(* IEC 61131-3 sources: STAR-PLC-Agent/results/raw/codex_matrix_resume_20261114/codex_deepseek/SELF004/functional/attempt_0001, 1 file *)

(* ---- test_program.st ---- *)
PROGRAM PLC_PRG
VAR
 BenchStep : UDINT := 0;
 BenchCalls : UDINT := 0;
 BenchDone : BOOL := FALSE;
 BenchUut0 : FB_Task;
 BenchUut1 : FB_Task;
 BenchUut2 : FB_Task;
 BenchUut3 : FB_Task;
 BenchUut4 : FB_Task;
 BenchUut5 : FB_Task;
 BenchUut6 : FB_Task;
 BenchUut7 : FB_Task;
 BenchUut8 : FB_Task;
 TraceIn_Start : ARRAY[0..60] OF BOOL;
 TraceIn_Stop : ARRAY[0..60] OF BOOL;
 TraceIn_AtExit : ARRAY[0..60] OF BOOL;
 TraceIn_Jam : ARRAY[0..60] OF BOOL;
 TraceIn_Reset : ARRAY[0..60] OF BOOL;
 TraceOut_Belt : ARRAY[0..60] OF BOOL;
 TraceOut_Complete : ARRAY[0..60] OF BOOL;
 TraceOut_Fault : ARRAY[0..60] OF BOOL;
END_VAR

IF NOT BenchDone THEN
 CASE BenchStep OF
 0:
   BenchUut0.Start := TRUE;
   BenchUut0.Stop := FALSE;
   BenchUut0.AtExit := FALSE;
   BenchUut0.Jam := FALSE;
   BenchUut0.Reset := FALSE;
   TraceIn_Start[0] := BenchUut0.Start;
   TraceIn_Stop[0] := BenchUut0.Stop;
   TraceIn_AtExit[0] := BenchUut0.AtExit;
   TraceIn_Jam[0] := BenchUut0.Jam;
   TraceIn_Reset[0] := BenchUut0.Reset;
   BenchUut0();
   TraceOut_Belt[0] := BenchUut0.Belt;
   TraceOut_Complete[0] := BenchUut0.Complete;
   TraceOut_Fault[0] := BenchUut0.Fault;
   BenchCalls := BenchCalls + 1;
 1:
   BenchUut0.Start := FALSE;
   BenchUut0.Stop := FALSE;
   BenchUut0.AtExit := FALSE;
   BenchUut0.Jam := FALSE;
   BenchUut0.Reset := FALSE;
   TraceIn_Start[1] := BenchUut0.Start;
   TraceIn_Stop[1] := BenchUut0.Stop;
   TraceIn_AtExit[1] := BenchUut0.AtExit;
   TraceIn_Jam[1] := BenchUut0.Jam;
   TraceIn_Reset[1] := BenchUut0.Reset;
   BenchUut0();
   TraceOut_Belt[1] := BenchUut0.Belt;
   TraceOut_Complete[1] := BenchUut0.Complete;
   TraceOut_Fault[1] := BenchUut0.Fault;
   BenchCalls := BenchCalls + 1;
 2:
   BenchUut0.Start := FALSE;
   BenchUut0.Stop := FALSE;
   BenchUut0.AtExit := TRUE;
   BenchUut0.Jam := FALSE;
   BenchUut0.Reset := FALSE;
   TraceIn_Start[2] := BenchUut0.Start;
   TraceIn_Stop[2] := BenchUut0.Stop;
   TraceIn_AtExit[2] := BenchUut0.AtExit;
   TraceIn_Jam[2] := BenchUut0.Jam;
   TraceIn_Reset[2] := BenchUut0.Reset;
   BenchUut0();
   TraceOut_Belt[2] := BenchUut0.Belt;
   TraceOut_Complete[2] := BenchUut0.Complete;
   TraceOut_Fault[2] := BenchUut0.Fault;
   BenchCalls := BenchCalls + 1;
 3:
   BenchUut0.Start := TRUE;
   BenchUut0.Stop := FALSE;
   BenchUut0.AtExit := FALSE;
   BenchUut0.Jam := FALSE;
   BenchUut0.Reset := FALSE;
   TraceIn_Start[3] := BenchUut0.Start;
   TraceIn_Stop[3] := BenchUut0.Stop;
   TraceIn_AtExit[3] := BenchUut0.AtExit;
   TraceIn_Jam[3] := BenchUut0.Jam;
   TraceIn_Reset[3] := BenchUut0.Reset;
   BenchUut0();
   TraceOut_Belt[3] := BenchUut0.Belt;
   TraceOut_Complete[3] := BenchUut0.Complete;
   TraceOut_Fault[3] := BenchUut0.Fault;
   BenchCalls := BenchCalls + 1;
 4:
   BenchUut0.Start := FALSE;
   BenchUut0.Stop := FALSE;
   BenchUut0.AtExit := FALSE;
   BenchUut0.Jam := FALSE;
   BenchUut0.Reset := TRUE;
   TraceIn_Start[4] := BenchUut0.Start;
   TraceIn_Stop[4] := BenchUut0.Stop;
   TraceIn_AtExit[4] := BenchUut0.AtExit;
   TraceIn_Jam[4] := BenchUut0.Jam;
   TraceIn_Reset[4] := BenchUut0.Reset;
   BenchUut0();
   TraceOut_Belt[4] := BenchUut0.Belt;
   TraceOut_Complete[4] := BenchUut0.Complete;
   TraceOut_Fault[4] := BenchUut0.Fault;
   BenchCalls := BenchCalls + 1;
 5:
   BenchUut1.Start := TRUE;
   BenchUut1.Stop := FALSE;
   BenchUut1.AtExit := FALSE;
   BenchUut1.Jam := FALSE;
   BenchUut1.Reset := FALSE;
   TraceIn_Start[5] := BenchUut1.Start;
   TraceIn_Stop[5] := BenchUut1.Stop;
   TraceIn_AtExit[5] := BenchUut1.AtExit;
   TraceIn_Jam[5] := BenchUut1.Jam;
   TraceIn_Reset[5] := BenchUut1.Reset;
   BenchUut1();
   TraceOut_Belt[5] := BenchUut1.Belt;
   TraceOut_Complete[5] := BenchUut1.Complete;
   TraceOut_Fault[5] := BenchUut1.Fault;
   BenchCalls := BenchCalls + 1;
 6:
   BenchUut1.Start := TRUE;
   BenchUut1.Stop := FALSE;
   BenchUut1.AtExit := FALSE;
   BenchUut1.Jam := TRUE;
   BenchUut1.Reset := TRUE;
   TraceIn_Start[6] := BenchUut1.Start;
   TraceIn_Stop[6] := BenchUut1.Stop;
   TraceIn_AtExit[6] := BenchUut1.AtExit;
   TraceIn_Jam[6] := BenchUut1.Jam;
   TraceIn_Reset[6] := BenchUut1.Reset;
   BenchUut1();
   TraceOut_Belt[6] := BenchUut1.Belt;
   TraceOut_Complete[6] := BenchUut1.Complete;
   TraceOut_Fault[6] := BenchUut1.Fault;
   BenchCalls := BenchCalls + 1;
 7:
   BenchUut1.Start := TRUE;
   BenchUut1.Stop := FALSE;
   BenchUut1.AtExit := FALSE;
   BenchUut1.Jam := FALSE;
   BenchUut1.Reset := FALSE;
   TraceIn_Start[7] := BenchUut1.Start;
   TraceIn_Stop[7] := BenchUut1.Stop;
   TraceIn_AtExit[7] := BenchUut1.AtExit;
   TraceIn_Jam[7] := BenchUut1.Jam;
   TraceIn_Reset[7] := BenchUut1.Reset;
   BenchUut1();
   TraceOut_Belt[7] := BenchUut1.Belt;
   TraceOut_Complete[7] := BenchUut1.Complete;
   TraceOut_Fault[7] := BenchUut1.Fault;
   BenchCalls := BenchCalls + 1;
 8:
   BenchUut1.Start := TRUE;
   BenchUut1.Stop := FALSE;
   BenchUut1.AtExit := FALSE;
   BenchUut1.Jam := FALSE;
   BenchUut1.Reset := TRUE;
   TraceIn_Start[8] := BenchUut1.Start;
   TraceIn_Stop[8] := BenchUut1.Stop;
   TraceIn_AtExit[8] := BenchUut1.AtExit;
   TraceIn_Jam[8] := BenchUut1.Jam;
   TraceIn_Reset[8] := BenchUut1.Reset;
   BenchUut1();
   TraceOut_Belt[8] := BenchUut1.Belt;
   TraceOut_Complete[8] := BenchUut1.Complete;
   TraceOut_Fault[8] := BenchUut1.Fault;
   BenchCalls := BenchCalls + 1;
 9:
   BenchUut1.Start := TRUE;
   BenchUut1.Stop := FALSE;
   BenchUut1.AtExit := TRUE;
   BenchUut1.Jam := FALSE;
   BenchUut1.Reset := FALSE;
   TraceIn_Start[9] := BenchUut1.Start;
   TraceIn_Stop[9] := BenchUut1.Stop;
   TraceIn_AtExit[9] := BenchUut1.AtExit;
   TraceIn_Jam[9] := BenchUut1.Jam;
   TraceIn_Reset[9] := BenchUut1.Reset;
   BenchUut1();
   TraceOut_Belt[9] := BenchUut1.Belt;
   TraceOut_Complete[9] := BenchUut1.Complete;
   TraceOut_Fault[9] := BenchUut1.Fault;
   BenchCalls := BenchCalls + 1;
 10:
   BenchUut1.Start := TRUE;
   BenchUut1.Stop := TRUE;
   BenchUut1.AtExit := FALSE;
   BenchUut1.Jam := FALSE;
   BenchUut1.Reset := FALSE;
   TraceIn_Start[10] := BenchUut1.Start;
   TraceIn_Stop[10] := BenchUut1.Stop;
   TraceIn_AtExit[10] := BenchUut1.AtExit;
   TraceIn_Jam[10] := BenchUut1.Jam;
   TraceIn_Reset[10] := BenchUut1.Reset;
   BenchUut1();
   TraceOut_Belt[10] := BenchUut1.Belt;
   TraceOut_Complete[10] := BenchUut1.Complete;
   TraceOut_Fault[10] := BenchUut1.Fault;
   BenchCalls := BenchCalls + 1;
 11:
   BenchUut2.Start := TRUE;
   BenchUut2.Stop := FALSE;
   BenchUut2.AtExit := FALSE;
   BenchUut2.Jam := FALSE;
   BenchUut2.Reset := FALSE;
   TraceIn_Start[11] := BenchUut2.Start;
   TraceIn_Stop[11] := BenchUut2.Stop;
   TraceIn_AtExit[11] := BenchUut2.AtExit;
   TraceIn_Jam[11] := BenchUut2.Jam;
   TraceIn_Reset[11] := BenchUut2.Reset;
   BenchUut2();
   TraceOut_Belt[11] := BenchUut2.Belt;
   TraceOut_Complete[11] := BenchUut2.Complete;
   TraceOut_Fault[11] := BenchUut2.Fault;
   BenchCalls := BenchCalls + 1;
 12:
   BenchUut2.Start := FALSE;
   BenchUut2.Stop := TRUE;
   BenchUut2.AtExit := TRUE;
   BenchUut2.Jam := FALSE;
   BenchUut2.Reset := FALSE;
   TraceIn_Start[12] := BenchUut2.Start;
   TraceIn_Stop[12] := BenchUut2.Stop;
   TraceIn_AtExit[12] := BenchUut2.AtExit;
   TraceIn_Jam[12] := BenchUut2.Jam;
   TraceIn_Reset[12] := BenchUut2.Reset;
   BenchUut2();
   TraceOut_Belt[12] := BenchUut2.Belt;
   TraceOut_Complete[12] := BenchUut2.Complete;
   TraceOut_Fault[12] := BenchUut2.Fault;
   BenchCalls := BenchCalls + 1;
 13:
   BenchUut2.Start := TRUE;
   BenchUut2.Stop := FALSE;
   BenchUut2.AtExit := FALSE;
   BenchUut2.Jam := FALSE;
   BenchUut2.Reset := FALSE;
   TraceIn_Start[13] := BenchUut2.Start;
   TraceIn_Stop[13] := BenchUut2.Stop;
   TraceIn_AtExit[13] := BenchUut2.AtExit;
   TraceIn_Jam[13] := BenchUut2.Jam;
   TraceIn_Reset[13] := BenchUut2.Reset;
   BenchUut2();
   TraceOut_Belt[13] := BenchUut2.Belt;
   TraceOut_Complete[13] := BenchUut2.Complete;
   TraceOut_Fault[13] := BenchUut2.Fault;
   BenchCalls := BenchCalls + 1;
 14:
   BenchUut2.Start := FALSE;
   BenchUut2.Stop := FALSE;
   BenchUut2.AtExit := FALSE;
   BenchUut2.Jam := FALSE;
   BenchUut2.Reset := TRUE;
   TraceIn_Start[14] := BenchUut2.Start;
   TraceIn_Stop[14] := BenchUut2.Stop;
   TraceIn_AtExit[14] := BenchUut2.AtExit;
   TraceIn_Jam[14] := BenchUut2.Jam;
   TraceIn_Reset[14] := BenchUut2.Reset;
   BenchUut2();
   TraceOut_Belt[14] := BenchUut2.Belt;
   TraceOut_Complete[14] := BenchUut2.Complete;
   TraceOut_Fault[14] := BenchUut2.Fault;
   BenchCalls := BenchCalls + 1;
 15:
   BenchUut2.Start := TRUE;
   BenchUut2.Stop := FALSE;
   BenchUut2.AtExit := FALSE;
   BenchUut2.Jam := FALSE;
   BenchUut2.Reset := FALSE;
   TraceIn_Start[15] := BenchUut2.Start;
   TraceIn_Stop[15] := BenchUut2.Stop;
   TraceIn_AtExit[15] := BenchUut2.AtExit;
   TraceIn_Jam[15] := BenchUut2.Jam;
   TraceIn_Reset[15] := BenchUut2.Reset;
   BenchUut2();
   TraceOut_Belt[15] := BenchUut2.Belt;
   TraceOut_Complete[15] := BenchUut2.Complete;
   TraceOut_Fault[15] := BenchUut2.Fault;
   BenchCalls := BenchCalls + 1;
 16:
   BenchUut2.Start := FALSE;
   BenchUut2.Stop := FALSE;
   BenchUut2.AtExit := TRUE;
   BenchUut2.Jam := FALSE;
   BenchUut2.Reset := FALSE;
   TraceIn_Start[16] := BenchUut2.Start;
   TraceIn_Stop[16] := BenchUut2.Stop;
   TraceIn_AtExit[16] := BenchUut2.AtExit;
   TraceIn_Jam[16] := BenchUut2.Jam;
   TraceIn_Reset[16] := BenchUut2.Reset;
   BenchUut2();
   TraceOut_Belt[16] := BenchUut2.Belt;
   TraceOut_Complete[16] := BenchUut2.Complete;
   TraceOut_Fault[16] := BenchUut2.Fault;
   BenchCalls := BenchCalls + 1;
 17:
   BenchUut2.Start := FALSE;
   BenchUut2.Stop := TRUE;
   BenchUut2.AtExit := TRUE;
   BenchUut2.Jam := FALSE;
   BenchUut2.Reset := FALSE;
   TraceIn_Start[17] := BenchUut2.Start;
   TraceIn_Stop[17] := BenchUut2.Stop;
   TraceIn_AtExit[17] := BenchUut2.AtExit;
   TraceIn_Jam[17] := BenchUut2.Jam;
   TraceIn_Reset[17] := BenchUut2.Reset;
   BenchUut2();
   TraceOut_Belt[17] := BenchUut2.Belt;
   TraceOut_Complete[17] := BenchUut2.Complete;
   TraceOut_Fault[17] := BenchUut2.Fault;
   BenchCalls := BenchCalls + 1;
 18:
   BenchUut2.Start := FALSE;
   BenchUut2.Stop := FALSE;
   BenchUut2.AtExit := FALSE;
   BenchUut2.Jam := TRUE;
   BenchUut2.Reset := FALSE;
   TraceIn_Start[18] := BenchUut2.Start;
   TraceIn_Stop[18] := BenchUut2.Stop;
   TraceIn_AtExit[18] := BenchUut2.AtExit;
   TraceIn_Jam[18] := BenchUut2.Jam;
   TraceIn_Reset[18] := BenchUut2.Reset;
   BenchUut2();
   TraceOut_Belt[18] := BenchUut2.Belt;
   TraceOut_Complete[18] := BenchUut2.Complete;
   TraceOut_Fault[18] := BenchUut2.Fault;
   BenchCalls := BenchCalls + 1;
 19:
   BenchUut2.Start := TRUE;
   BenchUut2.Stop := TRUE;
   BenchUut2.AtExit := FALSE;
   BenchUut2.Jam := FALSE;
   BenchUut2.Reset := FALSE;
   TraceIn_Start[19] := BenchUut2.Start;
   TraceIn_Stop[19] := BenchUut2.Stop;
   TraceIn_AtExit[19] := BenchUut2.AtExit;
   TraceIn_Jam[19] := BenchUut2.Jam;
   TraceIn_Reset[19] := BenchUut2.Reset;
   BenchUut2();
   TraceOut_Belt[19] := BenchUut2.Belt;
   TraceOut_Complete[19] := BenchUut2.Complete;
   TraceOut_Fault[19] := BenchUut2.Fault;
   BenchCalls := BenchCalls + 1;
 20:
   BenchUut2.Start := FALSE;
   BenchUut2.Stop := FALSE;
   BenchUut2.AtExit := FALSE;
   BenchUut2.Jam := FALSE;
   BenchUut2.Reset := TRUE;
   TraceIn_Start[20] := BenchUut2.Start;
   TraceIn_Stop[20] := BenchUut2.Stop;
   TraceIn_AtExit[20] := BenchUut2.AtExit;
   TraceIn_Jam[20] := BenchUut2.Jam;
   TraceIn_Reset[20] := BenchUut2.Reset;
   BenchUut2();
   TraceOut_Belt[20] := BenchUut2.Belt;
   TraceOut_Complete[20] := BenchUut2.Complete;
   TraceOut_Fault[20] := BenchUut2.Fault;
   BenchCalls := BenchCalls + 1;
 21:
   BenchUut3.Start := TRUE;
   BenchUut3.Stop := FALSE;
   BenchUut3.AtExit := FALSE;
   BenchUut3.Jam := FALSE;
   BenchUut3.Reset := FALSE;
   TraceIn_Start[21] := BenchUut3.Start;
   TraceIn_Stop[21] := BenchUut3.Stop;
   TraceIn_AtExit[21] := BenchUut3.AtExit;
   TraceIn_Jam[21] := BenchUut3.Jam;
   TraceIn_Reset[21] := BenchUut3.Reset;
   BenchUut3();
   TraceOut_Belt[21] := BenchUut3.Belt;
   TraceOut_Complete[21] := BenchUut3.Complete;
   TraceOut_Fault[21] := BenchUut3.Fault;
   BenchCalls := BenchCalls + 1;
 22:
   BenchUut3.Start := FALSE;
   BenchUut3.Stop := FALSE;
   BenchUut3.AtExit := FALSE;
   BenchUut3.Jam := FALSE;
   BenchUut3.Reset := FALSE;
   TraceIn_Start[22] := BenchUut3.Start;
   TraceIn_Stop[22] := BenchUut3.Stop;
   TraceIn_AtExit[22] := BenchUut3.AtExit;
   TraceIn_Jam[22] := BenchUut3.Jam;
   TraceIn_Reset[22] := BenchUut3.Reset;
   BenchUut3();
   TraceOut_Belt[22] := BenchUut3.Belt;
   TraceOut_Complete[22] := BenchUut3.Complete;
   TraceOut_Fault[22] := BenchUut3.Fault;
   BenchCalls := BenchCalls + 1;
 23:
   BenchUut3.Start := FALSE;
   BenchUut3.Stop := FALSE;
   BenchUut3.AtExit := TRUE;
   BenchUut3.Jam := FALSE;
   BenchUut3.Reset := FALSE;
   TraceIn_Start[23] := BenchUut3.Start;
   TraceIn_Stop[23] := BenchUut3.Stop;
   TraceIn_AtExit[23] := BenchUut3.AtExit;
   TraceIn_Jam[23] := BenchUut3.Jam;
   TraceIn_Reset[23] := BenchUut3.Reset;
   BenchUut3();
   TraceOut_Belt[23] := BenchUut3.Belt;
   TraceOut_Complete[23] := BenchUut3.Complete;
   TraceOut_Fault[23] := BenchUut3.Fault;
   BenchCalls := BenchCalls + 1;
 24:
   BenchUut3.Start := TRUE;
   BenchUut3.Stop := FALSE;
   BenchUut3.AtExit := FALSE;
   BenchUut3.Jam := FALSE;
   BenchUut3.Reset := FALSE;
   TraceIn_Start[24] := BenchUut3.Start;
   TraceIn_Stop[24] := BenchUut3.Stop;
   TraceIn_AtExit[24] := BenchUut3.AtExit;
   TraceIn_Jam[24] := BenchUut3.Jam;
   TraceIn_Reset[24] := BenchUut3.Reset;
   BenchUut3();
   TraceOut_Belt[24] := BenchUut3.Belt;
   TraceOut_Complete[24] := BenchUut3.Complete;
   TraceOut_Fault[24] := BenchUut3.Fault;
   BenchCalls := BenchCalls + 1;
 25:
   BenchUut3.Start := FALSE;
   BenchUut3.Stop := FALSE;
   BenchUut3.AtExit := FALSE;
   BenchUut3.Jam := FALSE;
   BenchUut3.Reset := TRUE;
   TraceIn_Start[25] := BenchUut3.Start;
   TraceIn_Stop[25] := BenchUut3.Stop;
   TraceIn_AtExit[25] := BenchUut3.AtExit;
   TraceIn_Jam[25] := BenchUut3.Jam;
   TraceIn_Reset[25] := BenchUut3.Reset;
   BenchUut3();
   TraceOut_Belt[25] := BenchUut3.Belt;
   TraceOut_Complete[25] := BenchUut3.Complete;
   TraceOut_Fault[25] := BenchUut3.Fault;
   BenchCalls := BenchCalls + 1;
 26:
   BenchUut3.Start := TRUE;
   BenchUut3.Stop := FALSE;
   BenchUut3.AtExit := FALSE;
   BenchUut3.Jam := FALSE;
   BenchUut3.Reset := TRUE;
   TraceIn_Start[26] := BenchUut3.Start;
   TraceIn_Stop[26] := BenchUut3.Stop;
   TraceIn_AtExit[26] := BenchUut3.AtExit;
   TraceIn_Jam[26] := BenchUut3.Jam;
   TraceIn_Reset[26] := BenchUut3.Reset;
   BenchUut3();
   TraceOut_Belt[26] := BenchUut3.Belt;
   TraceOut_Complete[26] := BenchUut3.Complete;
   TraceOut_Fault[26] := BenchUut3.Fault;
   BenchCalls := BenchCalls + 1;
 27:
   BenchUut3.Start := TRUE;
   BenchUut3.Stop := FALSE;
   BenchUut3.AtExit := FALSE;
   BenchUut3.Jam := FALSE;
   BenchUut3.Reset := TRUE;
   TraceIn_Start[27] := BenchUut3.Start;
   TraceIn_Stop[27] := BenchUut3.Stop;
   TraceIn_AtExit[27] := BenchUut3.AtExit;
   TraceIn_Jam[27] := BenchUut3.Jam;
   TraceIn_Reset[27] := BenchUut3.Reset;
   BenchUut3();
   TraceOut_Belt[27] := BenchUut3.Belt;
   TraceOut_Complete[27] := BenchUut3.Complete;
   TraceOut_Fault[27] := BenchUut3.Fault;
   BenchCalls := BenchCalls + 1;
 28:
   BenchUut4.Start := TRUE;
   BenchUut4.Stop := FALSE;
   BenchUut4.AtExit := FALSE;
   BenchUut4.Jam := FALSE;
   BenchUut4.Reset := FALSE;
   TraceIn_Start[28] := BenchUut4.Start;
   TraceIn_Stop[28] := BenchUut4.Stop;
   TraceIn_AtExit[28] := BenchUut4.AtExit;
   TraceIn_Jam[28] := BenchUut4.Jam;
   TraceIn_Reset[28] := BenchUut4.Reset;
   BenchUut4();
   TraceOut_Belt[28] := BenchUut4.Belt;
   TraceOut_Complete[28] := BenchUut4.Complete;
   TraceOut_Fault[28] := BenchUut4.Fault;
   BenchCalls := BenchCalls + 1;
 29:
   BenchUut4.Start := FALSE;
   BenchUut4.Stop := FALSE;
   BenchUut4.AtExit := FALSE;
   BenchUut4.Jam := FALSE;
   BenchUut4.Reset := FALSE;
   TraceIn_Start[29] := BenchUut4.Start;
   TraceIn_Stop[29] := BenchUut4.Stop;
   TraceIn_AtExit[29] := BenchUut4.AtExit;
   TraceIn_Jam[29] := BenchUut4.Jam;
   TraceIn_Reset[29] := BenchUut4.Reset;
   BenchUut4();
   TraceOut_Belt[29] := BenchUut4.Belt;
   TraceOut_Complete[29] := BenchUut4.Complete;
   TraceOut_Fault[29] := BenchUut4.Fault;
   BenchCalls := BenchCalls + 1;
 30:
   BenchUut4.Start := FALSE;
   BenchUut4.Stop := FALSE;
   BenchUut4.AtExit := TRUE;
   BenchUut4.Jam := FALSE;
   BenchUut4.Reset := FALSE;
   TraceIn_Start[30] := BenchUut4.Start;
   TraceIn_Stop[30] := BenchUut4.Stop;
   TraceIn_AtExit[30] := BenchUut4.AtExit;
   TraceIn_Jam[30] := BenchUut4.Jam;
   TraceIn_Reset[30] := BenchUut4.Reset;
   BenchUut4();
   TraceOut_Belt[30] := BenchUut4.Belt;
   TraceOut_Complete[30] := BenchUut4.Complete;
   TraceOut_Fault[30] := BenchUut4.Fault;
   BenchCalls := BenchCalls + 1;
 31:
   BenchUut4.Start := TRUE;
   BenchUut4.Stop := FALSE;
   BenchUut4.AtExit := FALSE;
   BenchUut4.Jam := FALSE;
   BenchUut4.Reset := FALSE;
   TraceIn_Start[31] := BenchUut4.Start;
   TraceIn_Stop[31] := BenchUut4.Stop;
   TraceIn_AtExit[31] := BenchUut4.AtExit;
   TraceIn_Jam[31] := BenchUut4.Jam;
   TraceIn_Reset[31] := BenchUut4.Reset;
   BenchUut4();
   TraceOut_Belt[31] := BenchUut4.Belt;
   TraceOut_Complete[31] := BenchUut4.Complete;
   TraceOut_Fault[31] := BenchUut4.Fault;
   BenchCalls := BenchCalls + 1;
 32:
   BenchUut4.Start := FALSE;
   BenchUut4.Stop := FALSE;
   BenchUut4.AtExit := FALSE;
   BenchUut4.Jam := FALSE;
   BenchUut4.Reset := TRUE;
   TraceIn_Start[32] := BenchUut4.Start;
   TraceIn_Stop[32] := BenchUut4.Stop;
   TraceIn_AtExit[32] := BenchUut4.AtExit;
   TraceIn_Jam[32] := BenchUut4.Jam;
   TraceIn_Reset[32] := BenchUut4.Reset;
   BenchUut4();
   TraceOut_Belt[32] := BenchUut4.Belt;
   TraceOut_Complete[32] := BenchUut4.Complete;
   TraceOut_Fault[32] := BenchUut4.Fault;
   BenchCalls := BenchCalls + 1;
 33:
   BenchUut4.Start := FALSE;
   BenchUut4.Stop := TRUE;
   BenchUut4.AtExit := FALSE;
   BenchUut4.Jam := FALSE;
   BenchUut4.Reset := TRUE;
   TraceIn_Start[33] := BenchUut4.Start;
   TraceIn_Stop[33] := BenchUut4.Stop;
   TraceIn_AtExit[33] := BenchUut4.AtExit;
   TraceIn_Jam[33] := BenchUut4.Jam;
   TraceIn_Reset[33] := BenchUut4.Reset;
   BenchUut4();
   TraceOut_Belt[33] := BenchUut4.Belt;
   TraceOut_Complete[33] := BenchUut4.Complete;
   TraceOut_Fault[33] := BenchUut4.Fault;
   BenchCalls := BenchCalls + 1;
 34:
   BenchUut4.Start := FALSE;
   BenchUut4.Stop := TRUE;
   BenchUut4.AtExit := FALSE;
   BenchUut4.Jam := FALSE;
   BenchUut4.Reset := TRUE;
   TraceIn_Start[34] := BenchUut4.Start;
   TraceIn_Stop[34] := BenchUut4.Stop;
   TraceIn_AtExit[34] := BenchUut4.AtExit;
   TraceIn_Jam[34] := BenchUut4.Jam;
   TraceIn_Reset[34] := BenchUut4.Reset;
   BenchUut4();
   TraceOut_Belt[34] := BenchUut4.Belt;
   TraceOut_Complete[34] := BenchUut4.Complete;
   TraceOut_Fault[34] := BenchUut4.Fault;
   BenchCalls := BenchCalls + 1;
 35:
   BenchUut5.Start := TRUE;
   BenchUut5.Stop := FALSE;
   BenchUut5.AtExit := FALSE;
   BenchUut5.Jam := FALSE;
   BenchUut5.Reset := FALSE;
   TraceIn_Start[35] := BenchUut5.Start;
   TraceIn_Stop[35] := BenchUut5.Stop;
   TraceIn_AtExit[35] := BenchUut5.AtExit;
   TraceIn_Jam[35] := BenchUut5.Jam;
   TraceIn_Reset[35] := BenchUut5.Reset;
   BenchUut5();
   TraceOut_Belt[35] := BenchUut5.Belt;
   TraceOut_Complete[35] := BenchUut5.Complete;
   TraceOut_Fault[35] := BenchUut5.Fault;
   BenchCalls := BenchCalls + 1;
 36:
   BenchUut5.Start := FALSE;
   BenchUut5.Stop := FALSE;
   BenchUut5.AtExit := FALSE;
   BenchUut5.Jam := FALSE;
   BenchUut5.Reset := FALSE;
   TraceIn_Start[36] := BenchUut5.Start;
   TraceIn_Stop[36] := BenchUut5.Stop;
   TraceIn_AtExit[36] := BenchUut5.AtExit;
   TraceIn_Jam[36] := BenchUut5.Jam;
   TraceIn_Reset[36] := BenchUut5.Reset;
   BenchUut5();
   TraceOut_Belt[36] := BenchUut5.Belt;
   TraceOut_Complete[36] := BenchUut5.Complete;
   TraceOut_Fault[36] := BenchUut5.Fault;
   BenchCalls := BenchCalls + 1;
 37:
   BenchUut5.Start := FALSE;
   BenchUut5.Stop := FALSE;
   BenchUut5.AtExit := TRUE;
   BenchUut5.Jam := FALSE;
   BenchUut5.Reset := FALSE;
   TraceIn_Start[37] := BenchUut5.Start;
   TraceIn_Stop[37] := BenchUut5.Stop;
   TraceIn_AtExit[37] := BenchUut5.AtExit;
   TraceIn_Jam[37] := BenchUut5.Jam;
   TraceIn_Reset[37] := BenchUut5.Reset;
   BenchUut5();
   TraceOut_Belt[37] := BenchUut5.Belt;
   TraceOut_Complete[37] := BenchUut5.Complete;
   TraceOut_Fault[37] := BenchUut5.Fault;
   BenchCalls := BenchCalls + 1;
 38:
   BenchUut5.Start := TRUE;
   BenchUut5.Stop := FALSE;
   BenchUut5.AtExit := FALSE;
   BenchUut5.Jam := FALSE;
   BenchUut5.Reset := FALSE;
   TraceIn_Start[38] := BenchUut5.Start;
   TraceIn_Stop[38] := BenchUut5.Stop;
   TraceIn_AtExit[38] := BenchUut5.AtExit;
   TraceIn_Jam[38] := BenchUut5.Jam;
   TraceIn_Reset[38] := BenchUut5.Reset;
   BenchUut5();
   TraceOut_Belt[38] := BenchUut5.Belt;
   TraceOut_Complete[38] := BenchUut5.Complete;
   TraceOut_Fault[38] := BenchUut5.Fault;
   BenchCalls := BenchCalls + 1;
 39:
   BenchUut5.Start := FALSE;
   BenchUut5.Stop := FALSE;
   BenchUut5.AtExit := FALSE;
   BenchUut5.Jam := FALSE;
   BenchUut5.Reset := TRUE;
   TraceIn_Start[39] := BenchUut5.Start;
   TraceIn_Stop[39] := BenchUut5.Stop;
   TraceIn_AtExit[39] := BenchUut5.AtExit;
   TraceIn_Jam[39] := BenchUut5.Jam;
   TraceIn_Reset[39] := BenchUut5.Reset;
   BenchUut5();
   TraceOut_Belt[39] := BenchUut5.Belt;
   TraceOut_Complete[39] := BenchUut5.Complete;
   TraceOut_Fault[39] := BenchUut5.Fault;
   BenchCalls := BenchCalls + 1;
 40:
   BenchUut5.Start := FALSE;
   BenchUut5.Stop := FALSE;
   BenchUut5.AtExit := TRUE;
   BenchUut5.Jam := FALSE;
   BenchUut5.Reset := TRUE;
   TraceIn_Start[40] := BenchUut5.Start;
   TraceIn_Stop[40] := BenchUut5.Stop;
   TraceIn_AtExit[40] := BenchUut5.AtExit;
   TraceIn_Jam[40] := BenchUut5.Jam;
   TraceIn_Reset[40] := BenchUut5.Reset;
   BenchUut5();
   TraceOut_Belt[40] := BenchUut5.Belt;
   TraceOut_Complete[40] := BenchUut5.Complete;
   TraceOut_Fault[40] := BenchUut5.Fault;
   BenchCalls := BenchCalls + 1;
 41:
   BenchUut5.Start := FALSE;
   BenchUut5.Stop := FALSE;
   BenchUut5.AtExit := TRUE;
   BenchUut5.Jam := FALSE;
   BenchUut5.Reset := TRUE;
   TraceIn_Start[41] := BenchUut5.Start;
   TraceIn_Stop[41] := BenchUut5.Stop;
   TraceIn_AtExit[41] := BenchUut5.AtExit;
   TraceIn_Jam[41] := BenchUut5.Jam;
   TraceIn_Reset[41] := BenchUut5.Reset;
   BenchUut5();
   TraceOut_Belt[41] := BenchUut5.Belt;
   TraceOut_Complete[41] := BenchUut5.Complete;
   TraceOut_Fault[41] := BenchUut5.Fault;
   BenchCalls := BenchCalls + 1;
 42:
   BenchUut6.Start := TRUE;
   BenchUut6.Stop := FALSE;
   BenchUut6.AtExit := FALSE;
   BenchUut6.Jam := FALSE;
   BenchUut6.Reset := FALSE;
   TraceIn_Start[42] := BenchUut6.Start;
   TraceIn_Stop[42] := BenchUut6.Stop;
   TraceIn_AtExit[42] := BenchUut6.AtExit;
   TraceIn_Jam[42] := BenchUut6.Jam;
   TraceIn_Reset[42] := BenchUut6.Reset;
   BenchUut6();
   TraceOut_Belt[42] := BenchUut6.Belt;
   TraceOut_Complete[42] := BenchUut6.Complete;
   TraceOut_Fault[42] := BenchUut6.Fault;
   BenchCalls := BenchCalls + 1;
 43:
   BenchUut6.Start := FALSE;
   BenchUut6.Stop := FALSE;
   BenchUut6.AtExit := FALSE;
   BenchUut6.Jam := FALSE;
   BenchUut6.Reset := FALSE;
   TraceIn_Start[43] := BenchUut6.Start;
   TraceIn_Stop[43] := BenchUut6.Stop;
   TraceIn_AtExit[43] := BenchUut6.AtExit;
   TraceIn_Jam[43] := BenchUut6.Jam;
   TraceIn_Reset[43] := BenchUut6.Reset;
   BenchUut6();
   TraceOut_Belt[43] := BenchUut6.Belt;
   TraceOut_Complete[43] := BenchUut6.Complete;
   TraceOut_Fault[43] := BenchUut6.Fault;
   BenchCalls := BenchCalls + 1;
 44:
   BenchUut6.Start := FALSE;
   BenchUut6.Stop := FALSE;
   BenchUut6.AtExit := TRUE;
   BenchUut6.Jam := FALSE;
   BenchUut6.Reset := FALSE;
   TraceIn_Start[44] := BenchUut6.Start;
   TraceIn_Stop[44] := BenchUut6.Stop;
   TraceIn_AtExit[44] := BenchUut6.AtExit;
   TraceIn_Jam[44] := BenchUut6.Jam;
   TraceIn_Reset[44] := BenchUut6.Reset;
   BenchUut6();
   TraceOut_Belt[44] := BenchUut6.Belt;
   TraceOut_Complete[44] := BenchUut6.Complete;
   TraceOut_Fault[44] := BenchUut6.Fault;
   BenchCalls := BenchCalls + 1;
 45:
   BenchUut6.Start := TRUE;
   BenchUut6.Stop := FALSE;
   BenchUut6.AtExit := FALSE;
   BenchUut6.Jam := FALSE;
   BenchUut6.Reset := FALSE;
   TraceIn_Start[45] := BenchUut6.Start;
   TraceIn_Stop[45] := BenchUut6.Stop;
   TraceIn_AtExit[45] := BenchUut6.AtExit;
   TraceIn_Jam[45] := BenchUut6.Jam;
   TraceIn_Reset[45] := BenchUut6.Reset;
   BenchUut6();
   TraceOut_Belt[45] := BenchUut6.Belt;
   TraceOut_Complete[45] := BenchUut6.Complete;
   TraceOut_Fault[45] := BenchUut6.Fault;
   BenchCalls := BenchCalls + 1;
 46:
   BenchUut6.Start := FALSE;
   BenchUut6.Stop := FALSE;
   BenchUut6.AtExit := FALSE;
   BenchUut6.Jam := FALSE;
   BenchUut6.Reset := TRUE;
   TraceIn_Start[46] := BenchUut6.Start;
   TraceIn_Stop[46] := BenchUut6.Stop;
   TraceIn_AtExit[46] := BenchUut6.AtExit;
   TraceIn_Jam[46] := BenchUut6.Jam;
   TraceIn_Reset[46] := BenchUut6.Reset;
   BenchUut6();
   TraceOut_Belt[46] := BenchUut6.Belt;
   TraceOut_Complete[46] := BenchUut6.Complete;
   TraceOut_Fault[46] := BenchUut6.Fault;
   BenchCalls := BenchCalls + 1;
 47:
   BenchUut6.Start := FALSE;
   BenchUut6.Stop := FALSE;
   BenchUut6.AtExit := FALSE;
   BenchUut6.Jam := TRUE;
   BenchUut6.Reset := TRUE;
   TraceIn_Start[47] := BenchUut6.Start;
   TraceIn_Stop[47] := BenchUut6.Stop;
   TraceIn_AtExit[47] := BenchUut6.AtExit;
   TraceIn_Jam[47] := BenchUut6.Jam;
   TraceIn_Reset[47] := BenchUut6.Reset;
   BenchUut6();
   TraceOut_Belt[47] := BenchUut6.Belt;
   TraceOut_Complete[47] := BenchUut6.Complete;
   TraceOut_Fault[47] := BenchUut6.Fault;
   BenchCalls := BenchCalls + 1;
 48:
   BenchUut6.Start := FALSE;
   BenchUut6.Stop := FALSE;
   BenchUut6.AtExit := FALSE;
   BenchUut6.Jam := TRUE;
   BenchUut6.Reset := TRUE;
   TraceIn_Start[48] := BenchUut6.Start;
   TraceIn_Stop[48] := BenchUut6.Stop;
   TraceIn_AtExit[48] := BenchUut6.AtExit;
   TraceIn_Jam[48] := BenchUut6.Jam;
   TraceIn_Reset[48] := BenchUut6.Reset;
   BenchUut6();
   TraceOut_Belt[48] := BenchUut6.Belt;
   TraceOut_Complete[48] := BenchUut6.Complete;
   TraceOut_Fault[48] := BenchUut6.Fault;
   BenchCalls := BenchCalls + 1;
 49:
   BenchUut7.Start := TRUE;
   BenchUut7.Stop := FALSE;
   BenchUut7.AtExit := FALSE;
   BenchUut7.Jam := FALSE;
   BenchUut7.Reset := FALSE;
   TraceIn_Start[49] := BenchUut7.Start;
   TraceIn_Stop[49] := BenchUut7.Stop;
   TraceIn_AtExit[49] := BenchUut7.AtExit;
   TraceIn_Jam[49] := BenchUut7.Jam;
   TraceIn_Reset[49] := BenchUut7.Reset;
   BenchUut7();
   TraceOut_Belt[49] := BenchUut7.Belt;
   TraceOut_Complete[49] := BenchUut7.Complete;
   TraceOut_Fault[49] := BenchUut7.Fault;
   BenchCalls := BenchCalls + 1;
 50:
   BenchUut7.Start := FALSE;
   BenchUut7.Stop := FALSE;
   BenchUut7.AtExit := FALSE;
   BenchUut7.Jam := FALSE;
   BenchUut7.Reset := FALSE;
   TraceIn_Start[50] := BenchUut7.Start;
   TraceIn_Stop[50] := BenchUut7.Stop;
   TraceIn_AtExit[50] := BenchUut7.AtExit;
   TraceIn_Jam[50] := BenchUut7.Jam;
   TraceIn_Reset[50] := BenchUut7.Reset;
   BenchUut7();
   TraceOut_Belt[50] := BenchUut7.Belt;
   TraceOut_Complete[50] := BenchUut7.Complete;
   TraceOut_Fault[50] := BenchUut7.Fault;
   BenchCalls := BenchCalls + 1;
 51:
   BenchUut7.Start := FALSE;
   BenchUut7.Stop := FALSE;
   BenchUut7.AtExit := TRUE;
   BenchUut7.Jam := FALSE;
   BenchUut7.Reset := FALSE;
   TraceIn_Start[51] := BenchUut7.Start;
   TraceIn_Stop[51] := BenchUut7.Stop;
   TraceIn_AtExit[51] := BenchUut7.AtExit;
   TraceIn_Jam[51] := BenchUut7.Jam;
   TraceIn_Reset[51] := BenchUut7.Reset;
   BenchUut7();
   TraceOut_Belt[51] := BenchUut7.Belt;
   TraceOut_Complete[51] := BenchUut7.Complete;
   TraceOut_Fault[51] := BenchUut7.Fault;
   BenchCalls := BenchCalls + 1;
 52:
   BenchUut7.Start := TRUE;
   BenchUut7.Stop := FALSE;
   BenchUut7.AtExit := FALSE;
   BenchUut7.Jam := FALSE;
   BenchUut7.Reset := FALSE;
   TraceIn_Start[52] := BenchUut7.Start;
   TraceIn_Stop[52] := BenchUut7.Stop;
   TraceIn_AtExit[52] := BenchUut7.AtExit;
   TraceIn_Jam[52] := BenchUut7.Jam;
   TraceIn_Reset[52] := BenchUut7.Reset;
   BenchUut7();
   TraceOut_Belt[52] := BenchUut7.Belt;
   TraceOut_Complete[52] := BenchUut7.Complete;
   TraceOut_Fault[52] := BenchUut7.Fault;
   BenchCalls := BenchCalls + 1;
 53:
   BenchUut7.Start := FALSE;
   BenchUut7.Stop := FALSE;
   BenchUut7.AtExit := FALSE;
   BenchUut7.Jam := FALSE;
   BenchUut7.Reset := TRUE;
   TraceIn_Start[53] := BenchUut7.Start;
   TraceIn_Stop[53] := BenchUut7.Stop;
   TraceIn_AtExit[53] := BenchUut7.AtExit;
   TraceIn_Jam[53] := BenchUut7.Jam;
   TraceIn_Reset[53] := BenchUut7.Reset;
   BenchUut7();
   TraceOut_Belt[53] := BenchUut7.Belt;
   TraceOut_Complete[53] := BenchUut7.Complete;
   TraceOut_Fault[53] := BenchUut7.Fault;
   BenchCalls := BenchCalls + 1;
 54:
   BenchUut7.Start := FALSE;
   BenchUut7.Stop := FALSE;
   BenchUut7.AtExit := FALSE;
   BenchUut7.Jam := FALSE;
   BenchUut7.Reset := FALSE;
   TraceIn_Start[54] := BenchUut7.Start;
   TraceIn_Stop[54] := BenchUut7.Stop;
   TraceIn_AtExit[54] := BenchUut7.AtExit;
   TraceIn_Jam[54] := BenchUut7.Jam;
   TraceIn_Reset[54] := BenchUut7.Reset;
   BenchUut7();
   TraceOut_Belt[54] := BenchUut7.Belt;
   TraceOut_Complete[54] := BenchUut7.Complete;
   TraceOut_Fault[54] := BenchUut7.Fault;
   BenchCalls := BenchCalls + 1;
 55:
   BenchUut7.Start := FALSE;
   BenchUut7.Stop := FALSE;
   BenchUut7.AtExit := FALSE;
   BenchUut7.Jam := FALSE;
   BenchUut7.Reset := FALSE;
   TraceIn_Start[55] := BenchUut7.Start;
   TraceIn_Stop[55] := BenchUut7.Stop;
   TraceIn_AtExit[55] := BenchUut7.AtExit;
   TraceIn_Jam[55] := BenchUut7.Jam;
   TraceIn_Reset[55] := BenchUut7.Reset;
   BenchUut7();
   TraceOut_Belt[55] := BenchUut7.Belt;
   TraceOut_Complete[55] := BenchUut7.Complete;
   TraceOut_Fault[55] := BenchUut7.Fault;
   BenchCalls := BenchCalls + 1;
 56:
   BenchUut8.Start := TRUE;
   BenchUut8.Stop := FALSE;
   BenchUut8.AtExit := FALSE;
   BenchUut8.Jam := FALSE;
   BenchUut8.Reset := FALSE;
   TraceIn_Start[56] := BenchUut8.Start;
   TraceIn_Stop[56] := BenchUut8.Stop;
   TraceIn_AtExit[56] := BenchUut8.AtExit;
   TraceIn_Jam[56] := BenchUut8.Jam;
   TraceIn_Reset[56] := BenchUut8.Reset;
   BenchUut8();
   TraceOut_Belt[56] := BenchUut8.Belt;
   TraceOut_Complete[56] := BenchUut8.Complete;
   TraceOut_Fault[56] := BenchUut8.Fault;
   BenchCalls := BenchCalls + 1;
 57:
   BenchUut8.Start := TRUE;
   BenchUut8.Stop := TRUE;
   BenchUut8.AtExit := FALSE;
   BenchUut8.Jam := FALSE;
   BenchUut8.Reset := FALSE;
   TraceIn_Start[57] := BenchUut8.Start;
   TraceIn_Stop[57] := BenchUut8.Stop;
   TraceIn_AtExit[57] := BenchUut8.AtExit;
   TraceIn_Jam[57] := BenchUut8.Jam;
   TraceIn_Reset[57] := BenchUut8.Reset;
   BenchUut8();
   TraceOut_Belt[57] := BenchUut8.Belt;
   TraceOut_Complete[57] := BenchUut8.Complete;
   TraceOut_Fault[57] := BenchUut8.Fault;
   BenchCalls := BenchCalls + 1;
 58:
   BenchUut8.Start := TRUE;
   BenchUut8.Stop := FALSE;
   BenchUut8.AtExit := FALSE;
   BenchUut8.Jam := FALSE;
   BenchUut8.Reset := FALSE;
   TraceIn_Start[58] := BenchUut8.Start;
   TraceIn_Stop[58] := BenchUut8.Stop;
   TraceIn_AtExit[58] := BenchUut8.AtExit;
   TraceIn_Jam[58] := BenchUut8.Jam;
   TraceIn_Reset[58] := BenchUut8.Reset;
   BenchUut8();
   TraceOut_Belt[58] := BenchUut8.Belt;
   TraceOut_Complete[58] := BenchUut8.Complete;
   TraceOut_Fault[58] := BenchUut8.Fault;
   BenchCalls := BenchCalls + 1;
 59:
   BenchUut8.Start := TRUE;
   BenchUut8.Stop := FALSE;
   BenchUut8.AtExit := FALSE;
   BenchUut8.Jam := TRUE;
   BenchUut8.Reset := FALSE;
   TraceIn_Start[59] := BenchUut8.Start;
   TraceIn_Stop[59] := BenchUut8.Stop;
   TraceIn_AtExit[59] := BenchUut8.AtExit;
   TraceIn_Jam[59] := BenchUut8.Jam;
   TraceIn_Reset[59] := BenchUut8.Reset;
   BenchUut8();
   TraceOut_Belt[59] := BenchUut8.Belt;
   TraceOut_Complete[59] := BenchUut8.Complete;
   TraceOut_Fault[59] := BenchUut8.Fault;
   BenchCalls := BenchCalls + 1;
 60:
   BenchUut8.Start := TRUE;
   BenchUut8.Stop := TRUE;
   BenchUut8.AtExit := FALSE;
   BenchUut8.Jam := FALSE;
   BenchUut8.Reset := FALSE;
   TraceIn_Start[60] := BenchUut8.Start;
   TraceIn_Stop[60] := BenchUut8.Stop;
   TraceIn_AtExit[60] := BenchUut8.AtExit;
   TraceIn_Jam[60] := BenchUut8.Jam;
   TraceIn_Reset[60] := BenchUut8.Reset;
   BenchUut8();
   TraceOut_Belt[60] := BenchUut8.Belt;
   TraceOut_Complete[60] := BenchUut8.Complete;
   TraceOut_Fault[60] := BenchUut8.Fault;
   BenchCalls := BenchCalls + 1;
 END_CASE;
 BenchStep := BenchStep + 1;
 IF BenchStep >= 61 THEN BenchDone := TRUE; END_IF;
END_IF;
END_PROGRAM
